FUNCTION_BLOCK MultilineComment (* Erste Zeile des Kommentars zweite Zeile, die deutlich laenger ist als die erste und trotzdem komplett im Diagramm sichtbar sein muss, auch wenn sie breiter als das Netzwerk ist, denn dieser Text ist absichtlich laenger als die Mindestbreite des Netzwerks von 1112 Pixeln und erzwingt daher die Verbreiterung des Diagramms dritte Zeile *)
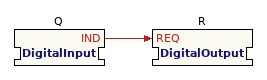
  FBS
    Q : DigitalInput;
    R : DigitalOutput;
  END_FBS
  EVENT_CONNECTIONS
    Q.IND TO R.REQ;
  END_CONNECTIONS
END_FUNCTION_BLOCK
